// TIA Portal V20 export
TYPE "Zylinder_v1_2"
   STRUCT
      Wartungsintervall : DInt;
      Fertigmeldung_Zylinder : Bool;
      Aktorzyklen : DInt;
      Auto_Frg_GS : Bool;
      Auto_Frg_AS : Bool;
      Manu_Frg_GS : Bool;
      Manu_Frg_AS : Bool;
      Richt_Frg_GS : Bool;
      Richt_Frg_AS : Bool;
      Status : Int;
   END_STRUCT;
END_TYPE
